(* IEC 61131-3 sources: RootPLC/conformance/cases/blocks (part 2) *)

(* ---- ok_rb_pump.st ---- *)
(* spec: [blocks.command] [blocks.interlock] [blocks.fault] [blocks.status]
   expect: ok
   libraries: RootBlocks *)
(* Test suite of RB_Pump (card blocks/cards/F04.PUMP.md). Every call passes
   the inputs that matter: block inputs keep their last value. *)
TEST pump_runs_like_a_motor
VAR p : RB_Pump; END_VAR
p(Mode := RB_MODE#Auto, AutoRun := TRUE, FbRunning := FALSE);
ASSERT_TRUE(p.Run);
ASSERT_FALSE(p.Running);
p(Mode := RB_MODE#Auto, AutoRun := TRUE, FbRunning := TRUE);
ASSERT_TRUE(p.Running);
ASSERT_EQ(UDINT#1, p.Status.Starts);
ASSERT_TRUE(p.Status.Commanded);
ASSERT_FALSE(p.Error);
p(Mode := RB_MODE#Manual, ManRun := FALSE, AutoRun := TRUE, FbRunning := TRUE);
ASSERT_FALSE(p.Run);
p(Mode := RB_MODE#Manual, ManRun := TRUE, Permissive := FALSE, FbRunning := FALSE);
ASSERT_FALSE(p.Run);
p(Mode := RB_MODE#Manual, ManRun := TRUE, Permissive := TRUE, Interlock := TRUE, FbRunning := FALSE);
ASSERT_FALSE(p.Run);
END_TEST

TEST pump_dry_run_trips_after_its_time
VAR p : RB_Pump; END_VAR
p(Mode := RB_MODE#Auto, AutoRun := TRUE, FbRunning := TRUE, DryRun := FALSE, DryRunTime := T#5s);
p(Mode := RB_MODE#Auto, AutoRun := TRUE, FbRunning := TRUE, DryRun := TRUE, DryRunTime := T#5s);
ADVANCE(T#4900ms);
p(Mode := RB_MODE#Auto, AutoRun := TRUE, FbRunning := TRUE, DryRun := TRUE, DryRunTime := T#5s);
ASSERT_FALSE(p.Error);
ASSERT_TRUE(p.Run);
ADVANCE(T#200ms);
p(Mode := RB_MODE#Auto, AutoRun := TRUE, FbRunning := TRUE, DryRun := TRUE, DryRunTime := T#5s);
ASSERT_TRUE(p.Error);
ASSERT_EQ(UDINT#4, p.ErrorID);
ASSERT_FALSE(p.Run);
ASSERT_TRUE(p.Status.Error);
ASSERT_EQ(UDINT#4, p.Status.ErrorID);
(* liquid back: still latched until reset *)
p(Mode := RB_MODE#Auto, AutoRun := TRUE, FbRunning := FALSE, DryRun := FALSE, DryRunTime := T#5s);
ASSERT_TRUE(p.Error);
ASSERT_FALSE(p.Run);
p(Mode := RB_MODE#Auto, AutoRun := TRUE, FbRunning := FALSE, DryRun := FALSE, DryRunTime := T#5s, Reset := TRUE);
ASSERT_FALSE(p.Error);
ASSERT_EQ(UDINT#0, p.ErrorID);
ASSERT_TRUE(p.Run);
END_TEST

TEST pump_dry_signal_while_stopped_is_no_fault
VAR p : RB_Pump; END_VAR
p(Mode := RB_MODE#Auto, AutoRun := FALSE, FbRunning := FALSE, DryRun := TRUE, DryRunTime := T#1s);
ADVANCE(T#5s);
p(Mode := RB_MODE#Auto, AutoRun := FALSE, FbRunning := FALSE, DryRun := TRUE, DryRunTime := T#1s);
ASSERT_FALSE(p.Error);
END_TEST

TEST pump_motor_faults_pass_through
VAR p : RB_Pump; q : RB_Pump; END_VAR
p(Mode := RB_MODE#Auto, AutoRun := TRUE, FbRunning := TRUE, Overload := TRUE);
ASSERT_TRUE(p.Error);
ASSERT_EQ(UDINT#3, p.ErrorID);
q(Mode := RB_MODE#Auto, AutoRun := TRUE, FbRunning := FALSE, FeedbackTime := T#1s, Feedback := TRUE);
ADVANCE(T#1100ms);
q(Mode := RB_MODE#Auto, AutoRun := TRUE, FbRunning := FALSE, FeedbackTime := T#1s, Feedback := TRUE);
ASSERT_EQ(UDINT#1, q.ErrorID);
ASSERT_TRUE(q.Error);
END_TEST

TEST pump_motor_fault_during_dry_running_wins
VAR p : RB_Pump; END_VAR
p(Mode := RB_MODE#Auto, AutoRun := TRUE, FbRunning := TRUE, DryRun := TRUE, DryRunTime := T#2s);
ADVANCE(T#1s);
p(Mode := RB_MODE#Auto, AutoRun := TRUE, FbRunning := TRUE, DryRun := TRUE, Overload := TRUE, DryRunTime := T#2s);
ASSERT_EQ(UDINT#3, p.ErrorID);
ADVANCE(T#2s);
p(Mode := RB_MODE#Auto, AutoRun := TRUE, FbRunning := FALSE, DryRun := TRUE, Overload := TRUE, DryRunTime := T#2s);
ASSERT_EQ(UDINT#3, p.ErrorID);
END_TEST

(* ---- ok_rb_round2.st ---- *)
(* spec: [blocks.mode] [blocks.interlock] [blocks.fault] [blocks.status] [blocks.testable]
   expect: ok
   libraries: RootBlocks *)
(* Test suites of RB_AnalogLimits (F08.LIMITS), RB_Ratio (F06.RATIO),
   RB_MotorTwoSpeed (F04.MOTOR.2SPEED), RB_Merge (F12.MERGE) and
   RB_Schedule (F03.SCHEDULE). Every call passes the inputs that matter:
   block inputs keep their last value. *)
TEST limits_with_hysteresis
VAR m : RB_AnalogLimits; END_VAR
m(Value := 50.0);
ASSERT_FALSE(m.HiHi OR m.Hi OR m.Lo OR m.LoLo OR m.Error);
m(Value := 85.0);
ASSERT_FALSE(m.Hi);
m(Value := 85.5);
ASSERT_TRUE(m.Hi);
ASSERT_FALSE(m.HiHi);
m(Value := 95.0);
ASSERT_FALSE(m.HiHi);
m(Value := 95.5);
ASSERT_TRUE(m.HiHi AND m.Hi);
(* back inside: active until Hysteresis below the limit *)
m(Value := 94.0);
ASSERT_TRUE(m.HiHi);
m(Value := 93.9);
ASSERT_FALSE(m.HiHi);
ASSERT_TRUE(m.Hi);
m(Value := 84.0);
ASSERT_TRUE(m.Hi);
m(Value := 83.9);
ASSERT_FALSE(m.Hi);
m(Value := 15.0);
ASSERT_FALSE(m.Lo);
m(Value := 14.5);
ASSERT_TRUE(m.Lo);
m(Value := 5.0);
ASSERT_FALSE(m.LoLo);
m(Value := 4.5);
ASSERT_TRUE(m.LoLo AND m.Lo);
m(Value := 6.0);
ASSERT_TRUE(m.LoLo);
m(Value := 6.1);
ASSERT_FALSE(m.LoLo);
m(Value := 16.0);
ASSERT_TRUE(m.Lo);
m(Value := 16.1);
ASSERT_FALSE(m.Lo);
END_TEST

TEST limits_enable_and_settings
VAR m : RB_AnalogLimits; END_VAR
m(Value := 99.0, EnHH := FALSE);
ASSERT_FALSE(m.HiHi);
ASSERT_TRUE(m.Hi);
m(EnH := FALSE);
ASSERT_FALSE(m.Hi);
m(Value := 1.0, EnLL := FALSE);
ASSERT_TRUE(m.Lo);
ASSERT_FALSE(m.LoLo);
m(EnL := FALSE);
ASSERT_FALSE(m.Lo);
(* limits out of order *)
m(Value := 99.0, EnHH := TRUE, EnH := TRUE, EnL := TRUE, EnLL := TRUE, H := 96.0);
ASSERT_TRUE(m.Error);
ASSERT_EQ(UDINT#1, m.ErrorID);
ASSERT_FALSE(m.HiHi OR m.Hi);
m(H := 95.0);
ASSERT_FALSE(m.Error);
ASSERT_EQ(UDINT#0, m.ErrorID);
ASSERT_TRUE(m.HiHi AND m.Hi);
m(Value := 0.0, L := 4.0);
ASSERT_TRUE(m.Error);
ASSERT_FALSE(m.Lo OR m.LoLo);
m(L := 5.0);
ASSERT_FALSE(m.Error);
ASSERT_TRUE(m.Lo AND m.LoLo);
m(L := 95.0);
ASSERT_TRUE(m.Error);
m(L := 15.0, Hysteresis := -1.0);
ASSERT_TRUE(m.Error);
m(Hysteresis := 0.0);
ASSERT_FALSE(m.Error);
END_TEST

TEST ratio_set_point
VAR r : RB_Ratio; END_VAR
r(Wild := 40.0, Ratio := 1.5, Bias := 2.0);
ASSERT_TRUE(ABS(r.SP - 62.0) < 0.001);
ASSERT_FALSE(r.Limited);
r(Wild := 80.0);
ASSERT_TRUE(ABS(r.SP - 100.0) < 0.001);
ASSERT_TRUE(r.Limited);
r(Wild := 100.0 / 1.5 - 2.0 / 1.5);
ASSERT_FALSE(r.Limited);
r(Wild := -10.0);
ASSERT_TRUE(ABS(r.SP) < 0.001);
ASSERT_TRUE(r.Limited);
r(Wild := 10.0, SPMin := 20.0);
ASSERT_TRUE(ABS(r.SP - 20.0) < 0.001);
ASSERT_TRUE(r.Limited);
ASSERT_FALSE(r.Error);
r(Wild := 12.0);
ASSERT_FALSE(r.Limited);
(* limits the wrong way round *)
r(SPMin := 60.0, SPMax := 50.0);
ASSERT_TRUE(r.Error);
ASSERT_EQ(UDINT#1, r.ErrorID);
ASSERT_TRUE(ABS(r.SP - 60.0) < 0.001);
ASSERT_TRUE(r.Limited);
r(SPMin := 50.0);
ASSERT_FALSE(r.Error);
ASSERT_EQ(UDINT#0, r.ErrorID);
END_TEST

TEST two_speed_motor_changes_speed_through_off
VAR m : RB_MotorTwoSpeed; END_VAR
m(Mode := RB_MODE#Auto, AutoRun := TRUE, AutoFast := FALSE);
ASSERT_TRUE(m.Slow);
ASSERT_FALSE(m.Fast);
ASSERT_FALSE(m.Running);
m(FbSlow := TRUE);
ASSERT_TRUE(m.Running);
ASSERT_FALSE(m.AtFast);
(* to fast: both off for Changeover first *)
m(AutoFast := TRUE, FbSlow := TRUE);
ASSERT_FALSE(m.Slow OR m.Fast);
ADVANCE(T#400ms);
m(FbSlow := FALSE);
ASSERT_FALSE(m.Slow OR m.Fast);
ADVANCE(T#100ms);
m();
ASSERT_TRUE(m.Fast);
ASSERT_FALSE(m.Slow);
ASSERT_FALSE(m.AtFast);
m(FbFast := TRUE);
ASSERT_TRUE(m.AtFast);
ASSERT_FALSE(m.Error);
ADVANCE(T#5s);
m();
ASSERT_TRUE(m.Fast);
(* back to slow, a request flipping during the gap is taken at its end *)
m(AutoFast := FALSE);
ASSERT_FALSE(m.Fast OR m.Slow);
ADVANCE(T#200ms);
m(AutoFast := TRUE, FbFast := FALSE);
ASSERT_FALSE(m.Fast OR m.Slow);
ADVANCE(T#300ms);
m();
ASSERT_TRUE(m.Fast);
(* stop; a start goes straight to the requested speed *)
m(AutoRun := FALSE);
ASSERT_FALSE(m.Fast OR m.Slow);
m(AutoRun := TRUE, AutoFast := FALSE, FbFast := FALSE, FbSlow := FALSE);
ASSERT_TRUE(m.Slow);
ASSERT_FALSE(m.Fast);
ASSERT_EQ(UDINT#2, m.Status.Starts);
END_TEST

TEST two_speed_motor_modes_and_faults
VAR m : RB_MotorTwoSpeed; END_VAR
m(Mode := RB_MODE#Manual, ManRun := TRUE, ManFast := TRUE, AutoRun := TRUE, AutoFast := FALSE);
ASSERT_TRUE(m.Fast);
m(Mode := RB_MODE#Off);
ASSERT_FALSE(m.Fast OR m.Slow);
m(Mode := RB_MODE#Auto, FbSlow := TRUE);
ASSERT_TRUE(m.Slow);
m(Overload := TRUE);
ASSERT_TRUE(m.Error);
ASSERT_EQ(UDINT#3, m.ErrorID);
ASSERT_FALSE(m.Fast OR m.Slow);
ASSERT_TRUE(m.Status.Error);
m(Overload := FALSE, Reset := TRUE);
ASSERT_FALSE(m.Error);
ASSERT_TRUE(m.Slow);
(* no feedback from either contactor *)
m(Reset := FALSE, FbSlow := FALSE, FeedbackTime := T#1s);
ADVANCE(T#1s);
m();
ASSERT_TRUE(m.Error);
ASSERT_EQ(UDINT#1, m.ErrorID);
m(Reset := TRUE, Feedback := FALSE, Interlock := TRUE);
ASSERT_FALSE(m.Slow);
m(Reset := FALSE, Interlock := FALSE, AutoRun := FALSE);
m(AutoRun := TRUE, Permissive := FALSE);
ASSERT_FALSE(m.Slow);
m(Permissive := TRUE, RestartDelay := T#1s);
ASSERT_FALSE(m.Slow);
ADVANCE(T#1s);
m();
ASSERT_TRUE(m.Slow);
ASSERT_TRUE(m.Running);
m(Changeover := T#1s, AutoFast := TRUE);
ADVANCE(T#900ms);
m();
ASSERT_FALSE(m.Fast);
ADVANCE(T#100ms);
m();
ASSERT_TRUE(m.Fast);
ASSERT_TRUE(m.AtFast);
END_TEST

TEST merge_alternates_and_counts
VAR g : RB_Merge; END_VAR
g(WaitingA := TRUE, WaitingB := TRUE, Clear := FALSE);
ASSERT_FALSE(g.ReleaseA OR g.ReleaseB);
g(Clear := TRUE);
ASSERT_TRUE(g.ReleaseA);
ASSERT_FALSE(g.ReleaseB);
(* the part passes the merge eye *)
g(MergeEye := TRUE);
ASSERT_TRUE(g.ReleaseA);
g(MergeEye := FALSE);
ASSERT_EQ(UDINT#1, g.FromA);
ASSERT_TRUE(g.ReleaseB);
ASSERT_FALSE(g.ReleaseA);
g(MergeEye := TRUE);
g(MergeEye := FALSE);
ASSERT_EQ(UDINT#1, g.FromB);
ASSERT_TRUE(g.ReleaseA);
g(MergeEye := TRUE);
g(MergeEye := FALSE, WaitingA := TRUE, WaitingB := FALSE);
ASSERT_EQ(UDINT#2, g.FromA);
(* only A waits: A again *)
ASSERT_TRUE(g.ReleaseA);
g(MergeEye := TRUE);
g(MergeEye := FALSE, WaitingA := FALSE, WaitingB := TRUE, Clear := FALSE);
ASSERT_FALSE(g.ReleaseA OR g.ReleaseB);
g(Clear := TRUE);
ASSERT_TRUE(g.ReleaseB);
(* an eye pulse with nothing released is not counted *)
g(MergeEye := TRUE);
g(MergeEye := FALSE, WaitingB := FALSE);
g(MergeEye := TRUE);
g(MergeEye := FALSE);
ASSERT_EQ(UDINT#3, g.FromA);
ASSERT_EQ(UDINT#2, g.FromB);
ASSERT_FALSE(g.ReleaseA OR g.ReleaseB);
END_TEST

TEST merge_priority_and_timeout
VAR g : RB_Merge; END_VAR
g(WaitingA := TRUE, WaitingB := TRUE, Clear := TRUE, PriorityA := TRUE, Timeout := T#2s);
ASSERT_TRUE(g.ReleaseA);
g(MergeEye := TRUE);
g(MergeEye := FALSE);
ASSERT_TRUE(g.ReleaseA);
(* nothing arrives at the eye *)
ADVANCE(T#1900ms);
g();
ASSERT_FALSE(g.Error);
ADVANCE(T#100ms);
g();
ASSERT_TRUE(g.Error);
ASSERT_EQ(UDINT#1, g.ErrorID);
ASSERT_FALSE(g.ReleaseA OR g.ReleaseB);
g(Reset := TRUE);
ASSERT_FALSE(g.Error);
ASSERT_EQ(UDINT#0, g.ErrorID);
ASSERT_TRUE(g.ReleaseA);
g(Reset := FALSE, PriorityA := FALSE);
g(MergeEye := TRUE);
g(MergeEye := FALSE);
ASSERT_TRUE(g.ReleaseB);
(* back-to-back releases: each one has its own Timeout *)
ADVANCE(T#1500ms);
g(MergeEye := TRUE);
g(MergeEye := FALSE);
ASSERT_TRUE(g.ReleaseA);
ADVANCE(T#1500ms);
g();
ASSERT_FALSE(g.Error);
ASSERT_TRUE(g.ReleaseA);
END_TEST

TEST schedule_day_window
VAR s : RB_Schedule; END_VAR
s(Now := TOD#05:59:59, Day := 1);
ASSERT_FALSE(s.Out);
s(Now := TOD#06:00:00);
ASSERT_TRUE(s.Out);
s(Now := TOD#21:59:59);
ASSERT_TRUE(s.Out);
s(Now := TOD#22:00:00);
ASSERT_FALSE(s.Out);
(* weekdays only *)
s(Now := TOD#12:00:00, Day := 6, Days := BYTE#16#1F);
ASSERT_FALSE(s.Out);
s(Day := 5);
ASSERT_TRUE(s.Out);
s(Day := 7, Days := BYTE#16#40);
ASSERT_TRUE(s.Out);
s(Enable := FALSE);
ASSERT_FALSE(s.Out);
s(Enable := TRUE, OnTime := TOD#12:00:00, OffTime := TOD#12:00:00);
ASSERT_FALSE(s.Out);
END_TEST

TEST schedule_overnight_and_errors
VAR s : RB_Schedule; END_VAR
(* a night shift Monday 22:00 to Tuesday 06:00, Mondays only *)
s(OnTime := TOD#22:00:00, OffTime := TOD#06:00:00, Days := BYTE#16#01, Now := TOD#21:00:00, Day := 1);
ASSERT_FALSE(s.Out);
s(Now := TOD#22:00:00);
ASSERT_TRUE(s.Out);
s(Now := TOD#05:00:00, Day := 2);
ASSERT_TRUE(s.Out);
s(Now := TOD#06:00:00);
ASSERT_FALSE(s.Out);
s(Now := TOD#23:00:00);
ASSERT_FALSE(s.Out);
s(Now := TOD#05:00:00, Day := 1);
ASSERT_FALSE(s.Out);
(* every day: the window ends exactly at OffTime *)
s(Days := BYTE#16#7F, Now := TOD#06:00:00, Day := 3);
ASSERT_FALSE(s.Out);
s(Now := TOD#21:59:59);
ASSERT_FALSE(s.Out);
(* Sunday night into Monday *)
s(Days := BYTE#16#40, Now := TOD#01:00:00, Day := 1);
ASSERT_TRUE(s.Out);
s(Day := 0);
ASSERT_TRUE(s.Error);
ASSERT_EQ(UDINT#1, s.ErrorID);
ASSERT_FALSE(s.Out);
s(Day := 8);
ASSERT_TRUE(s.Error);
s(Day := 7, Now := TOD#23:00:00);
ASSERT_FALSE(s.Error);
ASSERT_EQ(UDINT#0, s.ErrorID);
ASSERT_TRUE(s.Out);
END_TEST

(* ---- ok_rb_round3.st ---- *)
(* spec: [blocks.mode] [blocks.fault] [blocks.testable]
   expect: ok
   libraries: RootBlocks *)
(* Test suites of RB_Cascade (F06.CASCADE), RB_DutyStandby (F04.GROUP),
   RB_Totalizer (F09.TOTAL) and RB_OEE (F09.OEE). Every call passes the
   inputs that matter: block inputs keep their last value. *)
TEST cascade_modes
VAR c : RB_Cascade; END_VAR
c(Mode := RB_MODE#Off, SP := 70.0, PV := 60.0, InnerSP := 50.0, InnerPV := 40.0,
  KpInner := 2.0, ManValue := 33.0, OutMin := 5.0);
ASSERT_TRUE(ABS(c.Out - 5.0) < 0.001);
ASSERT_FALSE(c.InCascade);
c(Mode := RB_MODE#Manual);
ASSERT_TRUE(ABS(c.Out - 33.0) < 0.001);
(* set-point tracking: the inner set point follows the inner PV *)
ASSERT_TRUE(ABS(c.InnerSPUsed - 40.0) < 0.001);
ASSERT_FALSE(c.Saturated);
(* the inner loop alone on its own set point *)
c(Mode := RB_MODE#Auto, Cascade := FALSE);
ASSERT_FALSE(c.InCascade);
ASSERT_TRUE(ABS(c.InnerSPUsed - 50.0) < 0.001);
ASSERT_TRUE(ABS(c.Out - 20.0) < 0.001);
(* cascade: the outer loop sets the inner set point *)
c(Cascade := TRUE, KpOuter := 1.5);
ASSERT_TRUE(c.InCascade);
ASSERT_TRUE(ABS(c.InnerSPUsed - 15.0) < 0.001);
ASSERT_TRUE(ABS(c.Out - 5.0) < 0.001);
ASSERT_TRUE(c.Saturated);
c(SP := 200.0);
ASSERT_TRUE(ABS(c.InnerSPUsed - 100.0) < 0.001);
c(InnerSPMax := 80.0);
ASSERT_TRUE(ABS(c.InnerSPUsed - 80.0) < 0.001);
c(SP := 0.0, InnerSPMin := 10.0);
ASSERT_TRUE(ABS(c.InnerSPUsed - 10.0) < 0.001);
ASSERT_FALSE(c.Error);
ASSERT_EQ(UDINT#0, c.ErrorID);
END_TEST

TEST cascade_switches_bumpless
VAR c : RB_Cascade; END_VAR
(* in Manual the outer loop tracks the inner PV *)
c(Mode := RB_MODE#Manual, SP := 70.0, PV := 60.0, InnerPV := 40.0, KpOuter := 1.0,
  TiOuter := T#100s, KpInner := 1.0, TiInner := T#100s, ManValue := 30.0);
ADVANCE(T#100ms);
c();
c(Mode := RB_MODE#Auto);
ASSERT_TRUE(ABS(c.InnerSPUsed - 40.0) < 0.1);
ASSERT_TRUE(ABS(c.Out - 30.0) < 0.1);
(* then the outer integral moves the inner set point up *)
ADVANCE(T#10s);
c();
ASSERT_TRUE(c.InnerSPUsed > 40.5);
ASSERT_TRUE(c.Out > 30.0);
END_TEST

TEST cascade_errors
VAR c : RB_Cascade; END_VAR
c(Mode := RB_MODE#Auto, SP := 50.0, PV := 40.0, InnerPV := 40.0, OutMin := 100.0);
ASSERT_TRUE(c.Error);
ASSERT_EQ(UDINT#1, c.ErrorID);
ASSERT_TRUE(ABS(c.Out - 100.0) < 0.001);
c(OutMin := 0.0, Reset := TRUE);
ASSERT_FALSE(c.Error);
c(Reset := FALSE, InnerSPMin := 100.0);
ASSERT_TRUE(c.Error);
ASSERT_EQ(UDINT#11, c.ErrorID);
c(InnerSPMin := 0.0, Reset := TRUE);
ASSERT_FALSE(c.Error);
ASSERT_EQ(UDINT#0, c.ErrorID);
END_TEST

TEST duty_standby_least_hours_and_stages
VAR g : RB_DutyStandby; av : ARRAY[1..4] OF BOOL; h : ARRAY[1..4] OF REAL; k : INT; END_VAR
FOR k := 1 TO 4 DO av[k] := TRUE; END_FOR;
h[1] := 10.0; h[2] := 5.0; h[3] := 7.0; h[4] := 3.0;
g(Demand := 0, Available := av, Hours := h, StageDelay := T#5s);
ASSERT_EQ(0, g.Running);
ADVANCE(T#10s);
g(Demand := 1, Available := av, Hours := h);
ASSERT_TRUE(g.Run[4]);
ASSERT_EQ(1, g.Running);
ASSERT_FALSE(g.Shortfall);
(* the second unit waits for the stage delay, counted from the start *)
ADVANCE(T#100ms);
g(Demand := 2, Available := av, Hours := h);
ASSERT_EQ(1, g.Running);
ADVANCE(T#4800ms);
g(Demand := 2, Available := av, Hours := h);
ASSERT_EQ(1, g.Running);
ADVANCE(T#100ms);
g(Demand := 2, Available := av, Hours := h);
ASSERT_EQ(2, g.Running);
ASSERT_TRUE(g.Run[2]);
(* hours change while running: no swapping of running units *)
h[4] := 20.0;
ADVANCE(T#10s);
g(Demand := 2, Available := av, Hours := h);
ASSERT_TRUE(g.Run[4] AND g.Run[2]);
ASSERT_FALSE(g.Run[3]);
h[4] := 3.0;
(* unit 4 trips: replaced at once by the next with fewest hours *)
av[4] := FALSE;
g(Demand := 2, Available := av, Hours := h);
ASSERT_FALSE(g.Run[4]);
ASSERT_TRUE(g.Run[3]);
ASSERT_EQ(2, g.Running);
(* demand falls: the unit with the most hours stops *)
g(Demand := 1, Available := av, Hours := h);
ASSERT_FALSE(g.Run[3]);
ASSERT_TRUE(g.Run[2]);
ASSERT_EQ(1, g.Running);
g(Demand := 0, Available := av, Hours := h);
ASSERT_EQ(0, g.Running);
ASSERT_FALSE(g.Run[2]);
END_TEST

TEST duty_standby_shortfall_and_size
VAR g : RB_DutyStandby; av : ARRAY[1..4] OF BOOL; h : ARRAY[1..4] OF REAL; END_VAR
av[1] := TRUE; av[3] := TRUE;
h[1] := 2.0; h[3] := 1.0;
g(Demand := 3, Available := av, Hours := h);
ASSERT_TRUE(g.Run[3]);
ASSERT_TRUE(g.Shortfall);
g(Demand := 3, Available := av, Hours := h);
ASSERT_TRUE(g.Run[1]);
ASSERT_EQ(2, g.Running);
ASSERT_TRUE(g.Shortfall);
(* only two units fitted: unit 3 no longer counts *)
g(Demand := 3, Available := av, Hours := h, Used := 2);
ASSERT_FALSE(g.Run[3]);
ASSERT_TRUE(g.Run[1]);
ASSERT_EQ(1, g.Running);
ASSERT_TRUE(g.Shortfall);
av[2] := TRUE;
h[2] := 9.0;
g(Demand := 9, Available := av, Hours := h);
ASSERT_EQ(2, g.Running);
ASSERT_FALSE(g.Shortfall);
(* equal hours: the lowest number first *)
g(Demand := 0, Available := av, Hours := h, Used := 4);
h[1] := 1.0; h[2] := 1.0; h[3] := 1.0;
g(Demand := 1, Available := av, Hours := h);
ASSERT_TRUE(g.Run[1]);
(* equal hours: the lowest number stops first *)
g(Demand := 2, Available := av, Hours := h);
ASSERT_TRUE(g.Run[1] AND g.Run[2]);
g(Demand := 1, Available := av, Hours := h);
ASSERT_FALSE(g.Run[1]);
ASSERT_TRUE(g.Run[2]);
(* Used is limited to 1 .. 4 *)
g(Demand := 2, Available := av, Hours := h, Used := 0);
ASSERT_TRUE(g.Run[1]);
ASSERT_EQ(1, g.Running);
av[4] := TRUE;
g(Demand := 9, Available := av, Hours := h, Used := 9);
g(Demand := 9, Available := av, Hours := h, Used := 9);
g(Demand := 9, Available := av, Hours := h, Used := 9);
g(Demand := 9, Available := av, Hours := h, Used := 9);
ASSERT_EQ(4, g.Running);
END_TEST

TEST totalizer_counts_a_rate
VAR t : RB_Totalizer; END_VAR
t(Rate := 3600.0);
ASSERT_TRUE(ABS(t.Total) < 0.0001);
ADVANCE(T#1s);
t();
ASSERT_TRUE(ABS(t.Total - 1.0) < 0.0001);
ASSERT_TRUE(t.Counting);
ADVANCE(T#2s);
t(Hold := TRUE);
ASSERT_TRUE(ABS(t.Total - 1.0) < 0.0001);
ASSERT_FALSE(t.Counting);
(* the low-flow cut-off *)
ADVANCE(T#1s);
t(Hold := FALSE, LowCut := 3600.0);
ASSERT_TRUE(ABS(t.Total - 1.0) < 0.0001);
ADVANCE(T#1s);
t(Rate := 3601.0);
ASSERT_TRUE(t.Total > 1.9);
(* another time base: litres per minute *)
t(Reset := TRUE, LowCut := 0.0, Rate := 60.0, TimeBase := T#1m);
ASSERT_TRUE(ABS(t.Total) < 0.0001);
ADVANCE(T#3s);
t(Reset := FALSE);
ASSERT_TRUE(ABS(t.Total - 3.0) < 0.0001);
ADVANCE(T#1s);
t(TimeBase := T#0s);
ASSERT_FALSE(t.Counting);
ASSERT_TRUE(ABS(t.Total - 3.0) < 0.0001);
END_TEST

TEST totalizer_batch
VAR t : RB_Totalizer; END_VAR
t(Rate := 3600.0, Preset := 5.0);
ADVANCE(T#2s);
t();
ASSERT_TRUE(ABS(t.BatchTotal - 2.0) < 0.0001);
t(StartBatch := TRUE);
ASSERT_TRUE(ABS(t.BatchTotal) < 0.0001);
ASSERT_TRUE(ABS(t.Total - 2.0) < 0.0001);
ADVANCE(T#4s);
t(StartBatch := FALSE);
ASSERT_FALSE(t.BatchDone);
ADVANCE(T#1s);
t();
ASSERT_TRUE(t.BatchDone);
ASSERT_TRUE(ABS(t.BatchTotal - 5.0) < 0.0001);
t(StartBatch := TRUE);
ASSERT_FALSE(t.BatchDone);
(* without a preset the batch is never done *)
ADVANCE(T#10s);
t(StartBatch := FALSE, Preset := 0.0);
ASSERT_FALSE(t.BatchDone);
END_TEST

TEST oee_from_time_and_counts
VAR o : RB_OEE; i : INT; END_VAR
o(Planned := TRUE, Running := TRUE, IdealCycle := T#500ms);
ASSERT_TRUE(ABS(o.OEE) < 0.0001);
ASSERT_TRUE(ABS(o.Availability) < 0.0001);
FOR i := 1 TO 8 DO
    ADVANCE(T#1s);
    o(Good := i <= 6, Reject := i > 6);
    o(Good := FALSE, Reject := FALSE);
END_FOR;
FOR i := 1 TO 2 DO
    ADVANCE(T#1s);
    o(Running := FALSE);
END_FOR;
ASSERT_EQ(UDINT#6, o.GoodCount);
ASSERT_EQ(UDINT#2, o.RejectCount);
ASSERT_TRUE(ABS(o.PlannedTime - 10.0) < 0.001);
ASSERT_TRUE(ABS(o.RunTime - 8.0) < 0.001);
ASSERT_TRUE(ABS(o.Availability - 0.8) < 0.001);
ASSERT_TRUE(ABS(o.Performance - 0.5) < 0.001);
ASSERT_TRUE(ABS(o.Quality - 0.75) < 0.001);
ASSERT_TRUE(ABS(o.OEE - 0.3) < 0.001);
(* outside planned time nothing counts *)
ADVANCE(T#5s);
o(Planned := FALSE, Running := TRUE);
ASSERT_TRUE(ABS(o.PlannedTime - 10.0) < 0.001);
ASSERT_TRUE(ABS(o.RunTime - 8.0) < 0.001);
(* performance is at most 1 *)
o(IdealCycle := T#10s);
ASSERT_TRUE(ABS(o.Performance - 1.0) < 0.001);
o(Reset := TRUE);
ASSERT_EQ(UDINT#0, o.GoodCount);
ASSERT_EQ(UDINT#0, o.RejectCount);
ASSERT_TRUE(ABS(o.Performance) < 0.0001);
ASSERT_TRUE(ABS(o.Quality) < 0.0001);
ASSERT_TRUE(ABS(o.RunTime) < 0.0001);
END_TEST

TEST duty_standby_replaces_a_tripped_unit_at_once
VAR g : RB_DutyStandby; av : ARRAY[1..4] OF BOOL; h : ARRAY[1..4] OF REAL; END_VAR
av[1] := TRUE; av[2] := TRUE; av[3] := TRUE;
h[1] := 1.0; h[2] := 2.0; h[3] := 3.0;
g(Demand := 2, Available := av, Hours := h, StageDelay := T#5s, Used := 3);
ASSERT_TRUE(g.Run[1]);
ADVANCE(T#5s);
g(Demand := 2, Available := av, Hours := h);
ASSERT_TRUE(g.Run[2]);
(* one second after that start, unit 2 trips: unit 3 starts now *)
ADVANCE(T#1s);
av[2] := FALSE;
g(Demand := 2, Available := av, Hours := h);
ASSERT_FALSE(g.Run[2]);
ASSERT_TRUE(g.Run[3]);
ASSERT_EQ(2, g.Running);
END_TEST

(* ---- ok_rb_round5.st ---- *)
(* spec: [blocks.fault] [blocks.testable]
   expect: ok
   libraries: RootBlocks *)
(* Test suites of RB_Blink (F03.BLINK), RB_PWM (F06.PWM), RB_PulseRate
   (F01.PULSE), RB_ShiftTrack (F11.TRACK), RB_Vote2oo3 (F01.VOTE) and
   RB_Bypass (F02.BYPASS). Every call passes the inputs that matter: block
   inputs keep their last value. *)
TEST blink_on_and_off
VAR b : RB_Blink; END_VAR
b(Enable := FALSE);
ASSERT_FALSE(b.Out);
ASSERT_EQ(UDINT#0, b.Pulses);
b(Enable := TRUE);
ASSERT_TRUE(b.Out);
ASSERT_EQ(UDINT#1, b.Pulses);
ADVANCE(T#400ms);
b();
ASSERT_TRUE(b.Out);
ADVANCE(T#100ms);
b();
ASSERT_FALSE(b.Out);
ADVANCE(T#499ms);
b();
ASSERT_FALSE(b.Out);
ADVANCE(T#1ms);
b();
ASSERT_TRUE(b.Out);
ASSERT_EQ(UDINT#2, b.Pulses);
(* the phase is kept: a late call does not shift the next edge *)
ADVANCE(T#600ms);
b();
ASSERT_FALSE(b.Out);
ADVANCE(T#400ms);
b();
ASSERT_TRUE(b.Out);
ADVANCE(T#100ms);
b();
ASSERT_TRUE(b.Out);
(* off, then on again: starts on *)
b(Enable := FALSE);
ASSERT_FALSE(b.Out);
ADVANCE(T#250ms);
b(Enable := TRUE);
ASSERT_TRUE(b.Out);
ASSERT_EQ(UDINT#4, b.Pulses);
(* asymmetric *)
b(Enable := FALSE);
b(Enable := TRUE, OnTime := T#200ms, OffTime := T#800ms);
ADVANCE(T#200ms);
b();
ASSERT_FALSE(b.Out);
ADVANCE(T#700ms);
b();
ASSERT_FALSE(b.Out);
ADVANCE(T#100ms);
b();
ASSERT_TRUE(b.Out);
END_TEST

TEST pwm_duty_and_period
VAR p : RB_PWM; END_VAR
p(In := 25.0);
ASSERT_TRUE(p.Out);
ASSERT_EQ(T#500ms, p.OnTime);
ASSERT_FALSE(p.Error);
ADVANCE(T#400ms);
p();
ASSERT_TRUE(p.Out);
ADVANCE(T#100ms);
p();
ASSERT_FALSE(p.Out);
(* a new duty waits for the next period *)
ADVANCE(T#100ms);
p(In := 75.0);
ASSERT_FALSE(p.Out);
ASSERT_EQ(T#500ms, p.OnTime);
ADVANCE(T#1399ms);
p();
ASSERT_FALSE(p.Out);
ADVANCE(T#1ms);
p();
ASSERT_TRUE(p.Out);
ASSERT_EQ(T#1500ms, p.OnTime);
ADVANCE(T#1499ms);
p();
ASSERT_TRUE(p.Out);
ADVANCE(T#1ms);
p();
ASSERT_FALSE(p.Out);
(* disabled *)
p(Enable := FALSE);
ASSERT_FALSE(p.Out);
ASSERT_EQ(T#0s, p.OnTime);
p(Enable := TRUE, In := 0.0);
ASSERT_FALSE(p.Out);
p(Enable := FALSE);
p(Enable := TRUE, In := 150.0);
ASSERT_TRUE(p.Out);
ASSERT_EQ(T#2s, p.OnTime);
ADVANCE(T#1999ms);
p();
ASSERT_TRUE(p.Out);
END_TEST

TEST pwm_minimum_pulse_and_errors
VAR p : RB_PWM; END_VAR
p(In := 10.0, MinPulse := T#300ms);
ASSERT_EQ(T#0s, p.OnTime);
ASSERT_FALSE(p.Out);
p(Enable := FALSE);
p(Enable := TRUE, In := 90.0);
ASSERT_EQ(T#2s, p.OnTime);
p(Enable := FALSE);
p(Enable := TRUE, In := 15.0);
ASSERT_EQ(T#300ms, p.OnTime);
p(Enable := FALSE);
p(Enable := TRUE, In := 85.0);
ASSERT_EQ(T#1700ms, p.OnTime);
p(Period := T#0s);
ASSERT_TRUE(p.Error);
ASSERT_EQ(UDINT#1, p.ErrorID);
ASSERT_FALSE(p.Out);
p(Period := T#1s);
ASSERT_FALSE(p.Error);
ASSERT_EQ(UDINT#0, p.ErrorID);
ASSERT_TRUE(p.Out);
END_TEST

TEST pulse_rate_over_a_window
VAR r : RB_PulseRate; i : INT; END_VAR
r(Factor := 0.5);
FOR i := 1 TO 20 DO
    ADVANCE(T#50ms);
    r(Pulse := (i MOD 2) = 1);
END_FOR;
ASSERT_TRUE(ABS(r.Rate - 18000.0) < 0.001);
ASSERT_TRUE(ABS(r.Total - 5.0) < 0.0001);
ASSERT_EQ(UDINT#0, r.Pulses);
(* the next window, at half the pulse rate, per minute *)
FOR i := 1 TO 20 DO
    ADVANCE(T#50ms);
    r(Pulse := (i MOD 4) = 1, TimeBase := T#1m);
    IF i = 19 THEN
        ASSERT_EQ(UDINT#5, r.Pulses);
        ASSERT_TRUE(ABS(r.Rate - 18000.0) < 0.001);
    END_IF;
END_FOR;
ASSERT_TRUE(ABS(r.Rate - 150.0) < 0.001);
ASSERT_TRUE(ABS(r.Total - 7.5) < 0.0001);
(* no pulses: rate 0 after a window *)
ADVANCE(T#1s);
r(Pulse := FALSE);
ASSERT_TRUE(ABS(r.Rate) < 0.001);
r(Reset := TRUE);
ASSERT_TRUE(ABS(r.Total) < 0.0001);
r(Reset := FALSE, Window := T#0s, Pulse := TRUE);
ASSERT_TRUE(r.Error);
ASSERT_EQ(UDINT#1, r.ErrorID);
ASSERT_EQ(UDINT#0, r.Pulses);
r(Window := T#2s, Pulse := FALSE);
ASSERT_FALSE(r.Error);
ASSERT_EQ(UDINT#0, r.ErrorID);
END_TEST

TEST shift_track_moves_parts
VAR s : RB_ShiftTrack; i : INT; END_VAR
s(ReadPos := 3);
ASSERT_EQ(0, s.Occupied);
s(Shift := TRUE, InValue := 7);
ASSERT_EQ(DINT#7, s.Positions[1]);
s(Shift := FALSE);
s(Shift := TRUE, InValue := 0);
s(Shift := FALSE);
ASSERT_EQ(DINT#7, s.Positions[2]);
ASSERT_EQ(DINT#0, s.Positions[1]);
ASSERT_EQ(DINT#0, s.AtRead);
s(Shift := TRUE, InValue := 9);
ASSERT_EQ(DINT#7, s.AtRead);
ASSERT_EQ(2, s.Occupied);
(* the ejector takes it: removed there *)
s(Shift := FALSE, Remove := TRUE);
ASSERT_EQ(DINT#0, s.AtRead);
ASSERT_EQ(1, s.Occupied);
s(Remove := FALSE);
(* an entry falls out after position 64 *)
FOR i := 1 TO 63 DO
    s(Shift := TRUE, InValue := 0);
    s(Shift := FALSE);
END_FOR;
ASSERT_EQ(DINT#9, s.Positions[64]);
s(Shift := TRUE, InValue := 0);
ASSERT_EQ(0, s.Occupied);
s(Shift := FALSE, InValue := 5);
s(Shift := TRUE);
s(Shift := FALSE, ReadPos := 1);
ASSERT_EQ(DINT#5, s.AtRead);
s(Clear := TRUE);
ASSERT_EQ(0, s.Occupied);
ASSERT_EQ(DINT#0, s.AtRead);
END_TEST

TEST shift_track_read_position_range
VAR s : RB_ShiftTrack; END_VAR
s(Shift := TRUE, InValue := 4, ReadPos := 0);
ASSERT_TRUE(s.Error);
ASSERT_EQ(UDINT#1, s.ErrorID);
ASSERT_EQ(DINT#0, s.AtRead);
s(Shift := FALSE, ReadPos := 65, Remove := TRUE);
ASSERT_TRUE(s.Error);
ASSERT_EQ(1, s.Occupied);
s(ReadPos := 64, Remove := FALSE);
ASSERT_FALSE(s.Error);
ASSERT_EQ(UDINT#0, s.ErrorID);
s(ReadPos := 1);
ASSERT_EQ(DINT#4, s.AtRead);
END_TEST

TEST vote_median_average_and_deviation
VAR v : RB_Vote2oo3; END_VAR
v(A := 10.0, B := 11.0, C := 50.0);
ASSERT_TRUE(ABS(v.Value - 11.0) < 0.001);
ASSERT_EQ(3, v.Healthy);
ASSERT_FALSE(v.DevA OR v.DevB);
ASSERT_TRUE(v.DevC);
v(A := 50.0, B := 10.0, C := 11.0);
ASSERT_TRUE(ABS(v.Value - 11.0) < 0.001);
ASSERT_TRUE(v.DevA);
v(A := 11.0, B := 50.0, C := 10.0);
ASSERT_TRUE(ABS(v.Value - 11.0) < 0.001);
ASSERT_TRUE(v.DevB);
v(A := 10.0, B := 50.0, C := 11.0);
ASSERT_TRUE(ABS(v.Value - 11.0) < 0.001);
v(A := 11.0, B := 10.0, C := 50.0);
ASSERT_TRUE(ABS(v.Value - 11.0) < 0.001);
v(A := 50.0, B := 11.0, C := 10.0);
ASSERT_TRUE(ABS(v.Value - 11.0) < 0.001);
(* exactly MaxDev away is not a deviation *)
v(A := 9.0, B := 11.0, C := 13.0);
ASSERT_FALSE(v.DevA OR v.DevB OR v.DevC);
v(A := 11.0, B := 13.0, C := 9.0);
ASSERT_FALSE(v.DevA OR v.DevB OR v.DevC);
(* one unhealthy: the average of the other two *)
v(A := 10.0, B := 11.0, C := 50.0, OkC := FALSE);
ASSERT_TRUE(ABS(v.Value - 10.5) < 0.001);
ASSERT_EQ(2, v.Healthy);
ASSERT_FALSE(v.DevC);
v(OkC := TRUE, OkA := FALSE);
ASSERT_TRUE(ABS(v.Value - 30.5) < 0.001);
ASSERT_TRUE(v.DevB AND v.DevC);
ASSERT_FALSE(v.DevA);
v(OkA := TRUE, OkB := FALSE, A := 20.0, C := 22.0);
ASSERT_TRUE(ABS(v.Value - 21.0) < 0.001);
(* one left, then none: the last good value stays *)
v(OkA := FALSE);
ASSERT_TRUE(ABS(v.Value - 22.0) < 0.001);
ASSERT_EQ(1, v.Healthy);
ASSERT_FALSE(v.Error);
v(OkC := FALSE, C := 99.0);
ASSERT_TRUE(v.Error);
ASSERT_EQ(UDINT#1, v.ErrorID);
ASSERT_TRUE(ABS(v.Value - 22.0) < 0.001);
ASSERT_FALSE(v.DevA OR v.DevB OR v.DevC);
v(OkB := TRUE, B := 5.0);
ASSERT_FALSE(v.Error);
ASSERT_EQ(UDINT#0, v.ErrorID);
ASSERT_TRUE(ABS(v.Value - 5.0) < 0.001);
END_TEST

TEST bypass_with_key_and_time_limit
VAR y : RB_Bypass; END_VAR
y(Cond := FALSE, MaxTime := T#10s);
ASSERT_FALSE(y.Out);
(* no key: no bypass *)
y(Request := TRUE);
ASSERT_FALSE(y.Active);
y(Request := FALSE, Permit := TRUE);
y(Request := TRUE);
ASSERT_TRUE(y.Active);
ASSERT_TRUE(y.Out);
ASSERT_EQ(UDINT#1, y.Uses);
ASSERT_EQ(T#10s, y.Remaining);
ADVANCE(T#4s);
y(Request := FALSE);
ASSERT_EQ(T#6s, y.Remaining);
(* a second request while active changes nothing *)
y(Request := TRUE);
ASSERT_EQ(UDINT#1, y.Uses);
ADVANCE(T#6s);
y(Request := FALSE);
ASSERT_TRUE(y.Expired);
ASSERT_FALSE(y.Active);
ASSERT_FALSE(y.Out);
ASSERT_EQ(T#0s, y.Remaining);
y();
ASSERT_FALSE(y.Expired);
(* the condition itself still counts *)
y(Cond := TRUE);
ASSERT_TRUE(y.Out);
(* cancel, and the key turned back *)
y(Cond := FALSE, Request := TRUE);
ASSERT_TRUE(y.Active);
ASSERT_EQ(T#10s, y.Remaining);
y(Request := FALSE, Cancel := TRUE);
ASSERT_FALSE(y.Active);
y(Cancel := FALSE, Request := TRUE);
ASSERT_TRUE(y.Active);
ASSERT_EQ(UDINT#3, y.Uses);
y(Request := FALSE, Permit := FALSE);
ASSERT_FALSE(y.Active);
ASSERT_FALSE(y.Out);
END_TEST

(* ---- ok_rb_round6.st ---- *)
(* spec: [blocks.fault] [blocks.testable]
   expect: ok
   libraries: RootBlocks *)
(* Test suites of RB_SignalMonitor (F09.SIGNAL), RB_Trips (F02.TRIPS),
   RB_ZeroSpeed (F09.SPEED), RB_LevelSwitches (F12.LEVEL) and RB_EventLog
   (F08.EVENTS). Every call passes the inputs that matter: block inputs
   keep their last value. *)
TEST signal_monitor_stuck
VAR m : RB_SignalMonitor; i : INT; END_VAR
m(Value := 10.0, StuckTime := T#2s);
ASSERT_FALSE(m.Stuck);
ADVANCE(T#1900ms);
m();
ASSERT_FALSE(m.Stuck);
ADVANCE(T#100ms);
m();
ASSERT_TRUE(m.Stuck);
(* movement inside the band does not count *)
ADVANCE(T#1s);
m(Value := 10.05);
ASSERT_TRUE(m.Stuck);
m(Value := 10.2);
ASSERT_FALSE(m.Stuck);
(* a slow drift counts from where it last moved, not from call to call *)
FOR i := 1 TO 6 DO
    ADVANCE(T#1s);
    m(Value := 10.2 + INT_TO_REAL(i) * 0.06);
END_FOR;
ASSERT_FALSE(m.Stuck);
(* disabled: cleared, and a fresh start when enabled *)
ADVANCE(T#1500ms);
m();
m(Enable := FALSE);
ASSERT_FALSE(m.Stuck);
m(Enable := TRUE);
ADVANCE(T#1900ms);
m();
ASSERT_FALSE(m.Stuck);
(* exactly StuckBand is not a movement *)
m(Value := 0.0, StuckBand := 0.5, Enable := FALSE);
m(Enable := TRUE);
ADVANCE(T#1500ms);
m(Value := 0.5);
ADVANCE(T#500ms);
m(Value := 0.5);
ASSERT_TRUE(m.Stuck);
END_TEST

TEST signal_monitor_rate
VAR m : RB_SignalMonitor; END_VAR
m(Value := 0.0, MaxRate := 5.0);
ASSERT_TRUE(ABS(m.Rate) < 0.001);
ADVANCE(T#500ms);
m(Value := 2.5);
ASSERT_TRUE(ABS(m.Rate - 5.0) < 0.001);
ASSERT_FALSE(m.RateHigh);
ADVANCE(T#500ms);
m(Value := 5.5);
ASSERT_TRUE(ABS(m.Rate - 6.0) < 0.001);
ASSERT_TRUE(m.RateHigh);
ADVANCE(T#500ms);
m(Value := 2.0);
ASSERT_TRUE(ABS(m.Rate + 7.0) < 0.001);
ASSERT_TRUE(m.RateHigh);
(* two calls at the same instant keep the last rate *)
m(Value := 2.0);
ASSERT_TRUE(ABS(m.Rate + 7.0) < 0.001);
ADVANCE(T#500ms);
m(Value := 9.0, MaxRate := 0.0);
ASSERT_FALSE(m.RateHigh);
m(Enable := FALSE);
ASSERT_FALSE(m.RateHigh);
ASSERT_TRUE(ABS(m.Rate) < 0.001);
ADVANCE(T#100ms);
m(Enable := TRUE, MaxRate := 5.0, Value := 100.0);
ASSERT_TRUE(ABS(m.Rate) < 0.001);
ASSERT_FALSE(m.RateHigh);
END_TEST

TEST trips_latch_and_first_out
VAR t : RB_Trips; c : ARRAY[1..16] OF BOOL; END_VAR
t(Trip := c);
ASSERT_TRUE(t.Ok);
ASSERT_EQ(0, t.FirstOut);
c[4] := TRUE;
t(Trip := c);
ASSERT_FALSE(t.Ok);
ASSERT_EQ(WORD#16#0008, t.Latched);
ASSERT_EQ(4, t.FirstOut);
ASSERT_EQ(1, t.Active);
(* gone, but latched *)
c[4] := FALSE;
c[2] := TRUE;
t(Trip := c);
ASSERT_EQ(WORD#16#000A, t.Latched);
ASSERT_EQ(2, t.Active);
ASSERT_EQ(4, t.FirstOut);
(* reset clears only what has gone *)
t(Trip := c, Reset := TRUE);
ASSERT_EQ(WORD#16#0002, t.Latched);
ASSERT_EQ(4, t.FirstOut);
ASSERT_FALSE(t.Ok);
c[2] := FALSE;
t(Trip := c, Reset := FALSE);
ASSERT_FALSE(t.Ok);
t(Trip := c, Reset := TRUE);
ASSERT_TRUE(t.Ok);
ASSERT_EQ(0, t.FirstOut);
ASSERT_EQ(0, t.Active);
(* two in one call: the lowest is first *)
c[9] := TRUE;
c[7] := TRUE;
t(Trip := c, Reset := FALSE);
ASSERT_EQ(7, t.FirstOut);
END_TEST

TEST trips_unused
VAR t : RB_Trips; c : ARRAY[1..16] OF BOOL; END_VAR
c[16] := TRUE;
t(Trip := c, Used := WORD#16#7FFF);
ASSERT_TRUE(t.Ok);
t(Trip := c, Used := WORD#16#FFFF);
ASSERT_EQ(16, t.FirstOut);
ASSERT_EQ(WORD#16#8000, t.Latched);
(* taken out of use: no longer latched *)
c[16] := FALSE;
t(Trip := c, Used := WORD#16#7FFF);
ASSERT_TRUE(t.Ok);
c[1] := TRUE;
t(Trip := c);
ASSERT_EQ(1, t.FirstOut);
END_TEST

TEST zero_speed_monitor
VAR z : RB_ZeroSpeed; i : INT; END_VAR
z(Running := TRUE, Timeout := T#2s, StartDelay := T#5s);
ADVANCE(T#5s);
z();
ASSERT_TRUE(z.Monitoring);
ASSERT_FALSE(z.Error);
(* pulses every second keep it healthy *)
FOR i := 1 TO 10 DO
    ADVANCE(T#500ms);
    z(Pulse := TRUE);
    ADVANCE(T#500ms);
    z(Pulse := FALSE);
END_FOR;
ASSERT_FALSE(z.Error);
(* the gap counts from the last pulse edge, 500 ms ago *)
ADVANCE(T#1400ms);
z();
ASSERT_FALSE(z.Error);
ADVANCE(T#100ms);
z();
ASSERT_TRUE(z.Error);
ASSERT_EQ(UDINT#1, z.ErrorID);
(* latched until reset *)
z(Pulse := TRUE);
ASSERT_TRUE(z.Error);
z(Pulse := FALSE, Reset := TRUE);
ASSERT_FALSE(z.Error);
ASSERT_EQ(UDINT#0, z.ErrorID);
(* stopped: no monitoring; a restart waits StartDelay again *)
z(Reset := FALSE, Running := FALSE);
ASSERT_FALSE(z.Monitoring);
ADVANCE(T#10s);
z();
ASSERT_FALSE(z.Error);
z(Running := TRUE);
ADVANCE(T#4s);
z();
ASSERT_FALSE(z.Monitoring);
ASSERT_FALSE(z.Error);
ADVANCE(T#1s);
z();
ASSERT_TRUE(z.Monitoring);
ADVANCE(T#2s);
z();
ASSERT_TRUE(z.Error);
END_TEST

TEST level_switches_empty_a_sump
VAR l : RB_LevelSwitches; END_VAR
l();
ASSERT_FALSE(l.Pump);
ASSERT_TRUE(l.AlarmLow);
l(LowLowSw := TRUE, LowSw := TRUE);
ASSERT_FALSE(l.Pump);
ASSERT_FALSE(l.AlarmLow);
l(HighSw := TRUE);
ASSERT_TRUE(l.Pump);
l(HighSw := FALSE);
ASSERT_TRUE(l.Pump);
l(LowSw := FALSE);
ASSERT_FALSE(l.Pump);
(* high switch failed, high-high: the pump is forced on *)
l(LowSw := TRUE, HighHighSw := TRUE);
ASSERT_TRUE(l.Pump);
ASSERT_TRUE(l.AlarmHigh);
(* below low-low: never pump dry *)
l(HighHighSw := FALSE, HighSw := TRUE);
l(HighSw := FALSE, LowSw := TRUE, LowLowSw := FALSE);
ASSERT_FALSE(l.Pump);
ASSERT_TRUE(l.AlarmLow);
l(LowLowSw := TRUE);
ASSERT_TRUE(l.Pump);
(* disabled: off, and the demand is forgotten *)
l(Enable := FALSE);
ASSERT_FALSE(l.Pump);
l(Enable := TRUE);
ASSERT_FALSE(l.Pump);
END_TEST

TEST level_switches_fill_and_faults
VAR l : RB_LevelSwitches; END_VAR
l(Fill := TRUE, LowLowSw := TRUE, LowSw := FALSE);
ASSERT_TRUE(l.Pump);
l(LowSw := TRUE);
ASSERT_TRUE(l.Pump);
l(HighSw := TRUE);
ASSERT_FALSE(l.Pump);
l(HighSw := FALSE);
ASSERT_FALSE(l.Pump);
l(LowSw := FALSE);
ASSERT_TRUE(l.Pump);
l(HighHighSw := TRUE, LowSw := TRUE);
ASSERT_FALSE(l.Pump);
ASSERT_TRUE(l.AlarmHigh);
(* the pump runs too long *)
l(HighHighSw := FALSE, MaxRunTime := T#10s);
ASSERT_TRUE(l.Pump);
ADVANCE(T#9900ms);
l();
ASSERT_FALSE(l.Error);
ADVANCE(T#100ms);
l();
ASSERT_TRUE(l.Error);
ASSERT_EQ(UDINT#1, l.ErrorID);
ASSERT_FALSE(l.Pump);
l(Reset := TRUE, MaxRunTime := T#0s);
ASSERT_FALSE(l.Error);
ASSERT_EQ(UDINT#0, l.ErrorID);
ASSERT_TRUE(l.Pump);
ADVANCE(T#1h);
l(Reset := FALSE);
ASSERT_FALSE(l.Error);
(* contradicting switches *)
l(HighSw := TRUE, LowSw := FALSE);
ASSERT_TRUE(l.Error);
ASSERT_EQ(UDINT#2, l.ErrorID);
ASSERT_FALSE(l.Pump);
l(HighSw := FALSE, Reset := TRUE);
ASSERT_FALSE(l.Error);
END_TEST

TEST event_log_codes_and_stamps
VAR e : RB_EventLog; i : INT; END_VAR
e(Code := 101, Now := DT#2026-11-05-08:00:00);
ASSERT_EQ(0, e.Count);
e(Log := TRUE);
ASSERT_EQ(1, e.Count);
ASSERT_EQ(1, e.Newest);
ASSERT_EQ(DINT#101, e.Codes[1]);
ASSERT_TRUE(e.Stamps[1] = DT#2026-11-05-08:00:00);
e(Log := FALSE);
ASSERT_EQ(1, e.Count);
(* on change: each new non-zero code *)
e(OnChange := TRUE, Code := 5, Now := DT#2026-11-05-08:01:00);
ASSERT_EQ(2, e.Count);
ASSERT_TRUE(e.Stamps[2] = DT#2026-11-05-08:01:00);
e(Code := 5);
ASSERT_EQ(2, e.Count);
e(Code := 0);
ASSERT_EQ(2, e.Count);
e(Code := 5);
ASSERT_EQ(3, e.Count);
ASSERT_EQ(UDINT#3, e.Total);
(* without OnChange a change is not logged *)
e(OnChange := FALSE, Code := 7);
ASSERT_EQ(3, e.Count);
(* the ring keeps the last 32 *)
FOR i := 1 TO 37 DO
    e(Log := TRUE, Code := INT_TO_DINT(i));
    e(Log := FALSE);
END_FOR;
ASSERT_EQ(32, e.Count);
ASSERT_EQ(8, e.Newest);
ASSERT_EQ(DINT#37, e.Codes[8]);
ASSERT_EQ(UDINT#40, e.Total);
e(Clear := TRUE);
ASSERT_EQ(0, e.Count);
ASSERT_EQ(0, e.Newest);
e(Clear := FALSE, Log := TRUE);
ASSERT_EQ(1, e.Newest);
END_TEST

TEST peak_hold_minimum_maximum_average
VAR p : RB_PeakHold; END_VAR
p(Enable := FALSE, Value := 99.0);
ASSERT_EQ(UDINT#0, p.Samples);
ASSERT_TRUE(ABS(p.Maximum) < 0.001);
p(Enable := TRUE, Value := 4.0);
ASSERT_TRUE(ABS(p.Minimum - 4.0) < 0.001 AND ABS(p.Maximum - 4.0) < 0.001);
p(Value := 10.0);
p(Value := 1.0);
ASSERT_TRUE(ABS(p.Minimum - 1.0) < 0.001);
ASSERT_TRUE(ABS(p.Maximum - 10.0) < 0.001);
ASSERT_TRUE(ABS(p.Average - 5.0) < 0.001);
ASSERT_EQ(UDINT#3, p.Samples);
(* paused: nothing changes *)
p(Enable := FALSE, Value := 50.0);
ASSERT_TRUE(ABS(p.Maximum - 10.0) < 0.001);
ASSERT_EQ(UDINT#3, p.Samples);
(* reset: starts again from the next value *)
p(Reset := TRUE);
ASSERT_EQ(UDINT#0, p.Samples);
ASSERT_TRUE(ABS(p.Minimum) < 0.001 AND ABS(p.Maximum) < 0.001 AND ABS(p.Average) < 0.001);
p(Reset := FALSE, Enable := TRUE, Value := -3.0);
ASSERT_TRUE(ABS(p.Maximum + 3.0) < 0.001);
ASSERT_TRUE(ABS(p.Minimum + 3.0) < 0.001);
p(Reset := TRUE, Value := 7.0);
ASSERT_EQ(UDINT#1, p.Samples);
ASSERT_TRUE(ABS(p.Minimum - 7.0) < 0.001);
ASSERT_TRUE(ABS(p.Average - 7.0) < 0.001);
END_TEST

(* ---- ok_rb_scale.st ---- *)
(* spec: [blocks.library] [blocks.fault] [blocks.testable]
   expect: ok
   libraries: RootBlocks *)
(* Test suite of RB_Scale (card blocks/cards/F01.SCALE.md). *)
TEST scale_maps_linearly
VAR s : RB_Scale; END_VAR
s(Raw := 13824.0, RawMin := 0.0, RawMax := 27648.0, EngMin := 0.0, EngMax := 10.0);
ASSERT_TRUE(ABS(s.Value - 5.0) < 0.0001);
s(Raw := 4.0, RawMin := 4.0, RawMax := 20.0, EngMin := -50.0, EngMax := 150.0);
ASSERT_TRUE(ABS(s.Value + 50.0) < 0.0001);
s(Raw := 12.0, RawMin := 4.0, RawMax := 20.0, EngMin := -50.0, EngMax := 150.0);
ASSERT_TRUE(ABS(s.Value - 50.0) < 0.0001);
(* a falling characteristic *)
s(Raw := 0.0, RawMin := 0.0, RawMax := 100.0, EngMin := 10.0, EngMax := 0.0);
ASSERT_TRUE(ABS(s.Value - 10.0) < 0.0001);
ASSERT_FALSE(s.Error);
END_TEST

TEST scale_clamps_within_the_margin
VAR s : RB_Scale; END_VAR
s(Raw := 21.0, RawMin := 4.0, RawMax := 20.0, EngMin := 0.0, EngMax := 100.0, Margin := 2.0);
ASSERT_FALSE(s.Error);
ASSERT_TRUE(ABS(s.Value - 100.0) < 0.0001);
s(Raw := 3.0, RawMin := 4.0, RawMax := 20.0, EngMin := 0.0, EngMax := 100.0, Margin := 2.0);
ASSERT_TRUE(ABS(s.Value) < 0.0001);
s(Raw := 21.0, RawMin := 4.0, RawMax := 20.0, EngMin := 0.0, EngMax := 100.0, Margin := 2.0, Clamp := FALSE);
ASSERT_TRUE(ABS(s.Value - 106.25) < 0.0001);
(* a falling characteristic clamps too *)
s(Raw := 21.0, RawMin := 4.0, RawMax := 20.0, EngMin := 100.0, EngMax := 0.0, Margin := 2.0, Clamp := TRUE);
ASSERT_TRUE(ABS(s.Value) < 0.0001);
s(Raw := 3.0, RawMin := 4.0, RawMax := 20.0, EngMin := 100.0, EngMax := 0.0, Margin := 2.0);
ASSERT_TRUE(ABS(s.Value - 100.0) < 0.0001);
END_TEST

TEST scale_wire_break_latches_and_holds_the_last_value
VAR s : RB_Scale; END_VAR
s(Raw := 12.0, RawMin := 4.0, RawMax := 20.0, EngMin := 0.0, EngMax := 100.0, Margin := 0.5);
ASSERT_TRUE(ABS(s.Value - 50.0) < 0.0001);
s(Raw := 3.4, RawMin := 4.0, RawMax := 20.0, EngMin := 0.0, EngMax := 100.0, Margin := 0.5);
ASSERT_TRUE(s.Error);
ASSERT_EQ(UDINT#2, s.ErrorID);
ASSERT_TRUE(ABS(s.Value - 50.0) < 0.0001);
(* back in range: still latched, still the last valid value *)
s(Raw := 16.0, RawMin := 4.0, RawMax := 20.0, EngMin := 0.0, EngMax := 100.0, Margin := 0.5);
ASSERT_TRUE(s.Error);
ASSERT_TRUE(ABS(s.Value - 50.0) < 0.0001);
s(Raw := 16.0, RawMin := 4.0, RawMax := 20.0, EngMin := 0.0, EngMax := 100.0, Margin := 0.5, Reset := TRUE);
ASSERT_FALSE(s.Error);
ASSERT_EQ(UDINT#0, s.ErrorID);
ASSERT_TRUE(ABS(s.Value - 75.0) < 0.0001);
END_TEST

TEST scale_over_range_and_invalid_range
VAR s : RB_Scale; t : RB_Scale; END_VAR
s(Raw := 20.6, RawMin := 4.0, RawMax := 20.0, Margin := 0.5);
ASSERT_TRUE(s.Error);
ASSERT_EQ(UDINT#3, s.ErrorID);
s(Raw := 20.4, RawMin := 4.0, RawMax := 20.0, Margin := 0.5, Reset := TRUE);
ASSERT_FALSE(s.Error);
t(Raw := 5.0, RawMin := 4.0, RawMax := 4.0);
ASSERT_TRUE(t.Error);
ASSERT_EQ(UDINT#1, t.ErrorID);
(* the range may be given in either order *)
s(Raw := 4.2, RawMin := 20.0, RawMax := 4.0, EngMin := 0.0, EngMax := 100.0, Reset := FALSE);
ASSERT_FALSE(s.Error);
ASSERT_TRUE(ABS(s.Value - 98.75) < 0.0001);
END_TEST

TEST scale_limits_of_the_margin_are_valid
VAR s : RB_Scale; END_VAR
s(Raw := 20.5, RawMin := 4.0, RawMax := 20.0, Margin := 0.5);
ASSERT_FALSE(s.Error);
s(Raw := 3.5, RawMin := 4.0, RawMax := 20.0, Margin := 0.5);
ASSERT_FALSE(s.Error);
END_TEST

(* ---- ok_rb_signal.st ---- *)
(* spec: [blocks.testable] [blocks.library]
   expect: ok
   libraries: RootBlocks *)
(* Test suites of the S2 signal blocks: RB_CycleTime (F03.CYCLETIME),
   RB_FilterPT1 (F01.FILTER.PT1), RB_MovingAverage (F01.AVERAGE), RB_Ramp
   (F01.RAMP), RB_Deadband (F01.DEADBAND), RB_Debounce (F01.DEBOUNCE).
   Time comes from ADVANCE (the VM clock), as on a PLC. *)
TEST cycle_time_measures_seconds
VAR c : RB_CycleTime; END_VAR
c();
ASSERT_TRUE(c.FirstCall);
ASSERT_TRUE(ABS(c.Seconds) < 0.000001);
ASSERT_EQ(T#0s, c.Elapsed);
ADVANCE(T#250ms);
c();
ASSERT_FALSE(c.FirstCall);
ASSERT_TRUE(ABS(c.Seconds - 0.25) < 0.000001);
ASSERT_EQ(T#250ms, c.Elapsed);
ADVANCE(T#10ms);
c();
ASSERT_TRUE(ABS(c.Seconds - 0.01) < 0.000001);
c();
ASSERT_TRUE(ABS(c.Seconds) < 0.000001);
END_TEST

TEST cycle_time_survives_the_daily_restart
VAR c : RB_CycleTime; i : INT; total : LREAL; END_VAR
c();
FOR i := 1 TO 26 DO
    ADVANCE(T#1h);
    c();
    total := total + c.Seconds;
    ASSERT_EQ(T#1h, c.Elapsed);
END_FOR;
ASSERT_TRUE(ABS(total - 93600.0) < 0.001);
ASSERT_TRUE(ABS(c.Seconds - 3600.0) < 0.001);
END_TEST

TEST pt1_settles_with_its_time_constant
VAR f : RB_FilterPT1; i : INT; END_VAR
f(In := 10.0, T := T#1s);
ASSERT_TRUE(ABS(f.Out - 10.0) < 0.0001);
(* a step from 10 to 20: after one time constant about 63% of the step *)
FOR i := 1 TO 100 DO
    ADVANCE(T#10ms);
    f(In := 20.0, T := T#1s);
END_FOR;
ASSERT_TRUE(f.Out > 16.2 AND f.Out < 16.4);
FOR i := 1 TO 500 DO
    ADVANCE(T#10ms);
    f(In := 20.0, T := T#1s);
END_FOR;
ASSERT_TRUE(ABS(f.Out - 20.0) < 0.1);
(* falling as well *)
ADVANCE(T#1s);
f(In := 0.0, T := T#1s);
ASSERT_TRUE(f.Out > 9.9 AND f.Out < 10.1);
END_TEST

TEST pt1_track_and_zero_time_constant_pass_through
VAR f : RB_FilterPT1; g : RB_FilterPT1; END_VAR
f(In := 0.0, T := T#5s);
ADVANCE(T#100ms);
f(In := 50.0, T := T#5s, Track := TRUE);
ASSERT_TRUE(ABS(f.Out - 50.0) < 0.0001);
ADVANCE(T#100ms);
f(In := 0.0, T := T#5s, Track := FALSE);
ASSERT_TRUE(f.Out > 48.0 AND f.Out < 50.0);
g(In := 0.0, T := T#0s);
ADVANCE(T#100ms);
g(In := 7.0, T := T#0s);
ASSERT_TRUE(ABS(g.Out - 7.0) < 0.0001);
(* two calls at the same instant *)
g(In := 3.0, T := T#0s);
ASSERT_TRUE(ABS(g.Out - 3.0) < 0.0001);
END_TEST

TEST average_over_the_window
VAR a : RB_MovingAverage; END_VAR
a(In := 2.0, Window := 3);
ASSERT_TRUE(ABS(a.Out - 2.0) < 0.0001);
ASSERT_FALSE(a.Valid);
a(In := 4.0, Window := 3);
ASSERT_TRUE(ABS(a.Out - 3.0) < 0.0001);
a(In := 6.0, Window := 3);
ASSERT_TRUE(ABS(a.Out - 4.0) < 0.0001);
ASSERT_TRUE(a.Valid);
a(In := 8.0, Window := 3);
ASSERT_TRUE(ABS(a.Out - 6.0) < 0.0001);
a(In := 1.0, Window := 3, Reset := TRUE);
ASSERT_TRUE(ABS(a.Out - 1.0) < 0.0001);
ASSERT_FALSE(a.Valid);
END_TEST

TEST average_window_is_clamped
VAR a : RB_MovingAverage; b : RB_MovingAverage; i : INT; END_VAR
a(In := 5.0, Window := 0);
ASSERT_TRUE(a.Valid);
a(In := 9.0, Window := 0);
ASSERT_TRUE(ABS(a.Out - 9.0) < 0.0001);
FOR i := 1 TO 31 DO
    b(In := 1.0, Window := 40);
END_FOR;
ASSERT_FALSE(b.Valid);
b(In := 33.0, Window := 40);
ASSERT_TRUE(b.Valid);
ASSERT_TRUE(ABS(b.Out - 2.0) < 0.0001);
END_TEST

TEST ramp_limits_rise_and_fall
VAR r : RB_Ramp; i : INT; END_VAR
r(In := 0.0, RiseRate := 10.0, FallRate := 20.0);
ASSERT_TRUE(ABS(r.Out) < 0.0001);
ASSERT_FALSE(r.Busy);
ADVANCE(T#500ms);
r(In := 100.0, RiseRate := 10.0, FallRate := 20.0);
ASSERT_TRUE(ABS(r.Out - 5.0) < 0.001);
ASSERT_TRUE(r.Busy);
FOR i := 1 TO 20 DO
    ADVANCE(T#500ms);
    r(In := 100.0, RiseRate := 10.0, FallRate := 20.0);
END_FOR;
ASSERT_TRUE(ABS(r.Out - 100.0) < 0.001);
ASSERT_FALSE(r.Busy);
ADVANCE(T#1s);
r(In := 0.0, RiseRate := 10.0, FallRate := 20.0);
ASSERT_TRUE(ABS(r.Out - 80.0) < 0.001);
FOR i := 1 TO 10 DO
    ADVANCE(T#1s);
    r(In := 0.0, RiseRate := 10.0, FallRate := 20.0);
END_FOR;
ASSERT_TRUE(ABS(r.Out) < 0.001);
END_TEST

TEST ramp_rate_zero_and_track_pass_through
VAR r : RB_Ramp; END_VAR
r(In := 0.0, RiseRate := 0.0, FallRate := 5.0);
ADVANCE(T#100ms);
r(In := 40.0, RiseRate := 0.0, FallRate := 5.0);
ASSERT_TRUE(ABS(r.Out - 40.0) < 0.001);
ADVANCE(T#100ms);
r(In := 0.0, RiseRate := 0.0, FallRate := 5.0);
ASSERT_TRUE(ABS(r.Out - 39.5) < 0.001);
ADVANCE(T#100ms);
r(In := 0.0, RiseRate := 0.0, FallRate := 0.0);
ASSERT_TRUE(ABS(r.Out) < 0.001);
ADVANCE(T#100ms);
r(In := 60.0, RiseRate := 1.0, FallRate := 1.0, Track := TRUE);
ASSERT_TRUE(ABS(r.Out - 60.0) < 0.001);
END_TEST

TEST deadband_holds_until_the_input_moves_enough
VAR d : RB_Deadband; END_VAR
d(In := 10.0, Deadband := 0.5);
ASSERT_TRUE(ABS(d.Out - 10.0) < 0.0001);
d(In := 10.4, Deadband := 0.5);
ASSERT_TRUE(ABS(d.Out - 10.0) < 0.0001);
d(In := 9.5, Deadband := 0.5);
ASSERT_TRUE(ABS(d.Out - 10.0) < 0.0001);
d(In := 10.6, Deadband := 0.5);
ASSERT_TRUE(ABS(d.Out - 10.6) < 0.0001);
d(In := 10.2, Deadband := 0.5);
ASSERT_TRUE(ABS(d.Out - 10.6) < 0.0001);
d(In := 10.0, Deadband := 0.0);
ASSERT_TRUE(ABS(d.Out - 10.0) < 0.0001);
END_TEST

TEST debounce_needs_a_stable_contact
VAR b : RB_Debounce; END_VAR
b(In := TRUE, OnDelay := T#50ms, OffDelay := T#100ms);
ASSERT_FALSE(b.Out);
ADVANCE(T#40ms);
b(In := FALSE, OnDelay := T#50ms, OffDelay := T#100ms);
ADVANCE(T#20ms);
b(In := TRUE, OnDelay := T#50ms, OffDelay := T#100ms);
ADVANCE(T#40ms);
b(In := TRUE, OnDelay := T#50ms, OffDelay := T#100ms);
ASSERT_FALSE(b.Out);
ADVANCE(T#20ms);
b(In := TRUE, OnDelay := T#50ms, OffDelay := T#100ms);
ASSERT_TRUE(b.Out);
(* a short drop is ignored; a long one switches off *)
b(In := FALSE, OnDelay := T#50ms, OffDelay := T#100ms);
ADVANCE(T#90ms);
b(In := FALSE, OnDelay := T#50ms, OffDelay := T#100ms);
ASSERT_TRUE(b.Out);
b(In := TRUE, OnDelay := T#50ms, OffDelay := T#100ms);
b(In := FALSE, OnDelay := T#50ms, OffDelay := T#100ms);
ADVANCE(T#90ms);
b(In := FALSE, OnDelay := T#50ms, OffDelay := T#100ms);
ASSERT_TRUE(b.Out);
ADVANCE(T#20ms);
b(In := FALSE, OnDelay := T#50ms, OffDelay := T#100ms);
ASSERT_FALSE(b.Out);
END_TEST

(* ---- ok_rb_valve_onoff.st ---- *)
(* spec: [blocks.library] [blocks.command] [blocks.mode] [blocks.interlock] [blocks.fault] [blocks.feedback] [blocks.status] [blocks.testable]
   expect: ok
   libraries: RootBlocks *)
(* Test suite of RB_ValveOnOff (card blocks/cards/F04.VALVE.ONOFF.md). *)
TEST valve_auto_opens_and_reports
VAR v : RB_ValveOnOff; END_VAR
v(Mode := RB_MODE#Auto, AutoOpen := TRUE, FbOpen := FALSE, FbClosed := TRUE);
ASSERT_TRUE(v.Open);
ASSERT_FALSE(v.IsOpen);
ASSERT_TRUE(v.Status.Commanded);
ASSERT_FALSE(v.Status.Active);
v(Mode := RB_MODE#Auto, AutoOpen := TRUE, FbOpen := TRUE, FbClosed := FALSE);
ASSERT_TRUE(v.IsOpen);
ASSERT_FALSE(v.IsClosed);
ASSERT_TRUE(v.Status.Active);
ASSERT_EQ(UDINT#1, v.Status.Starts);
ASSERT_TRUE(v.Status.Mode = RB_MODE#Auto);
v(Mode := RB_MODE#Auto, AutoOpen := TRUE, FbOpen := TRUE, FbClosed := FALSE);
ASSERT_EQ(UDINT#1, v.Status.Starts);
v(Mode := RB_MODE#Auto, AutoOpen := FALSE, FbOpen := TRUE, FbClosed := FALSE);
ASSERT_FALSE(v.Open);
v(Mode := RB_MODE#Auto, AutoOpen := FALSE, FbOpen := FALSE, FbClosed := TRUE);
ASSERT_TRUE(v.IsClosed);
v(Mode := RB_MODE#Auto, AutoOpen := TRUE, FbOpen := FALSE, FbClosed := TRUE);
ASSERT_EQ(UDINT#2, v.Status.Starts);
ASSERT_FALSE(v.Error);
END_TEST

TEST valve_mode_selects_the_command
VAR v : RB_ValveOnOff; END_VAR
v(Mode := RB_MODE#Auto, ManOpen := TRUE, FbOpen := FALSE, FbClosed := TRUE);
ASSERT_FALSE(v.Open);
v(Mode := RB_MODE#Manual, ManOpen := TRUE, AutoOpen := FALSE, FbOpen := FALSE, FbClosed := TRUE);
ASSERT_TRUE(v.Open);
v(Mode := RB_MODE#Manual, ManOpen := FALSE, AutoOpen := TRUE, FbOpen := TRUE, FbClosed := FALSE);
ASSERT_FALSE(v.Open);
v(Mode := RB_MODE#Off, ManOpen := TRUE, AutoOpen := TRUE, FbOpen := FALSE, FbClosed := TRUE);
ASSERT_FALSE(v.Open);
ASSERT_TRUE(v.Status.Mode = RB_MODE#Off);
END_TEST

TEST valve_interlock_closes_in_every_mode
VAR v : RB_ValveOnOff; END_VAR
v(Mode := RB_MODE#Manual, ManOpen := TRUE, FbOpen := FALSE, FbClosed := TRUE);
v(Mode := RB_MODE#Manual, ManOpen := TRUE, FbOpen := TRUE, FbClosed := FALSE);
ASSERT_TRUE(v.Open);
v(Mode := RB_MODE#Manual, ManOpen := TRUE, Interlock := TRUE, FbOpen := TRUE, FbClosed := FALSE);
ASSERT_FALSE(v.Open);
v(Mode := RB_MODE#Auto, AutoOpen := TRUE, Interlock := TRUE, FbOpen := FALSE, FbClosed := TRUE);
ASSERT_FALSE(v.Open);
v(Mode := RB_MODE#Auto, AutoOpen := TRUE, Interlock := FALSE, FbOpen := FALSE, FbClosed := TRUE);
ASSERT_TRUE(v.Open);
END_TEST

TEST valve_permissive_is_needed_to_open_not_to_stay_open
VAR v : RB_ValveOnOff; END_VAR
v(Mode := RB_MODE#Auto, AutoOpen := TRUE, Permissive := FALSE, FbOpen := FALSE, FbClosed := TRUE);
ASSERT_FALSE(v.Open);
ASSERT_EQ(UDINT#0, v.Status.Starts);
v(Mode := RB_MODE#Auto, AutoOpen := TRUE, Permissive := TRUE, FbOpen := FALSE, FbClosed := TRUE);
ASSERT_TRUE(v.Open);
v(Mode := RB_MODE#Auto, AutoOpen := TRUE, Permissive := FALSE, FbOpen := TRUE, FbClosed := FALSE);
ASSERT_TRUE(v.Open);
END_TEST

TEST valve_does_not_open_in_time_latches_until_reset
VAR v : RB_ValveOnOff; END_VAR
(* stuck closed: the closed switch stays on *)
v(Mode := RB_MODE#Auto, AutoOpen := TRUE, FbOpen := FALSE, FbClosed := TRUE, FeedbackTime := T#2s);
ADVANCE(T#1900ms);
v(Mode := RB_MODE#Auto, AutoOpen := TRUE, FbOpen := FALSE, FbClosed := TRUE, FeedbackTime := T#2s);
ASSERT_FALSE(v.Error);
ADVANCE(T#200ms);
v(Mode := RB_MODE#Auto, AutoOpen := TRUE, FbOpen := FALSE, FbClosed := TRUE, FeedbackTime := T#2s);
ASSERT_TRUE(v.Error);
ASSERT_EQ(UDINT#1, v.ErrorID);
ASSERT_FALSE(v.Open);
ASSERT_TRUE(v.Status.Error);
ASSERT_EQ(UDINT#1, v.Status.ErrorID);
(* the cause goes away: the fault stays latched *)
ADVANCE(T#5s);
v(Mode := RB_MODE#Auto, AutoOpen := TRUE, FbOpen := FALSE, FbClosed := TRUE, FeedbackTime := T#2s);
ASSERT_TRUE(v.Error);
ASSERT_FALSE(v.Open);
(* reset: it opens again; still stuck, so the fault returns after 2 s *)
v(Mode := RB_MODE#Auto, AutoOpen := TRUE, FbOpen := FALSE, FbClosed := TRUE, FeedbackTime := T#2s, Reset := TRUE);
ASSERT_FALSE(v.Error);
ASSERT_EQ(UDINT#0, v.ErrorID);
ASSERT_TRUE(v.Open);
ADVANCE(T#2100ms);
v(Mode := RB_MODE#Auto, AutoOpen := TRUE, FbOpen := FALSE, FbClosed := TRUE, FeedbackTime := T#2s, Reset := TRUE);
ASSERT_TRUE(v.Error);
ASSERT_EQ(UDINT#1, v.ErrorID);
END_TEST

TEST valve_does_not_close_in_time
VAR v : RB_ValveOnOff; END_VAR
(* stuck open: no command, the open switch stays on *)
v(Mode := RB_MODE#Auto, FbOpen := TRUE, FeedbackTime := T#1s);
ADVANCE(T#1100ms);
v(Mode := RB_MODE#Auto, FbOpen := TRUE, FeedbackTime := T#1s);
ASSERT_TRUE(v.Error);
ASSERT_EQ(UDINT#2, v.ErrorID);
END_TEST

TEST valve_contradicting_feedback
VAR v : RB_ValveOnOff; END_VAR
v(Mode := RB_MODE#Auto, AutoOpen := TRUE, FbOpen := TRUE, FbClosed := TRUE, FeedbackTime := T#1s);
ADVANCE(T#900ms);
v(Mode := RB_MODE#Auto, AutoOpen := TRUE, FbOpen := TRUE, FbClosed := TRUE, FeedbackTime := T#1s);
ASSERT_FALSE(v.Error);
ADVANCE(T#200ms);
v(Mode := RB_MODE#Auto, AutoOpen := TRUE, FbOpen := TRUE, FbClosed := TRUE, FeedbackTime := T#1s);
ASSERT_TRUE(v.Error);
ASSERT_EQ(UDINT#3, v.ErrorID);
ASSERT_FALSE(v.IsOpen);
ASSERT_FALSE(v.IsClosed);
END_TEST

TEST valve_without_feedback_follows_the_command
VAR v : RB_ValveOnOff; END_VAR
v(Mode := RB_MODE#Auto, AutoOpen := TRUE, Feedback := FALSE, FeedbackTime := T#1s);
ASSERT_TRUE(v.IsOpen);
ASSERT_FALSE(v.IsClosed);
ADVANCE(T#5s);
v(Mode := RB_MODE#Auto, AutoOpen := TRUE, Feedback := FALSE, FeedbackTime := T#1s);
ASSERT_FALSE(v.Error);
v(Mode := RB_MODE#Auto, AutoOpen := FALSE, Feedback := FALSE, FeedbackTime := T#1s);
ASSERT_FALSE(v.IsOpen);
ASSERT_TRUE(v.IsClosed);
END_TEST

TEST valve_feedback_switched_on_starts_supervision_fresh
VAR v : RB_ValveOnOff; END_VAR
v(Mode := RB_MODE#Auto, AutoOpen := TRUE, Feedback := FALSE, FbOpen := FALSE, FbClosed := TRUE, FeedbackTime := T#1s);
ADVANCE(T#5s);
v(Mode := RB_MODE#Auto, AutoOpen := TRUE, Feedback := FALSE, FbOpen := FALSE, FbClosed := TRUE, FeedbackTime := T#1s);
v(Mode := RB_MODE#Auto, AutoOpen := TRUE, Feedback := TRUE, FbOpen := FALSE, FbClosed := TRUE, FeedbackTime := T#1s);
ASSERT_FALSE(v.Error);
ADVANCE(T#1100ms);
v(Mode := RB_MODE#Auto, AutoOpen := TRUE, Feedback := TRUE, FbOpen := FALSE, FbClosed := TRUE, FeedbackTime := T#1s);
ASSERT_TRUE(v.Error);
END_TEST

TEST valve_conflict_supervision_starts_fresh_too
VAR v : RB_ValveOnOff; END_VAR
v(Mode := RB_MODE#Auto, AutoOpen := TRUE, Feedback := FALSE, FbOpen := TRUE, FbClosed := TRUE, FeedbackTime := T#1s);
ADVANCE(T#5s);
v(Mode := RB_MODE#Auto, AutoOpen := TRUE, Feedback := FALSE, FbOpen := TRUE, FbClosed := TRUE, FeedbackTime := T#1s);
v(Mode := RB_MODE#Auto, AutoOpen := TRUE, Feedback := TRUE, FbOpen := TRUE, FbClosed := TRUE, FeedbackTime := T#1s);
ASSERT_FALSE(v.Error);
END_TEST
